PROGRAM MAIN
VAR
    fbMotionSystem : FB_MotionSystem;
    nState         : UDINT;
END_VAR

// Main program: start up the system, enable it, then run the exercise.
CASE nState OF
    0:  nState := 1;
    1:  IF fbMotionSystem.Startup() THEN
            nState := 30;
        END_IF
    30: IF fbMotionSystem.Starting(bReset := FALSE) THEN
            nState := 40;
        END_IF
    40: fbMotionSystem.Execute();   // drive in loops without stopping
END_CASE

fbMotionSystem.Cycle();

END_PROGRAM

(* stored: Version 1.1.0.1
   POU MAIN: Id {cafd9452-95b0-482f-a5bb-58f53d94daaf} *)
